Fanuc KAREL source: kt00743.KL

PROGRAM KT00743
%STACKSIZE=65535
%PRIORITY=65535
%NOLOCKGROUP
VAR
ARG : ARRAY[4] OF VECTOR
OUT : INTEGER
BEGIN
-- UNSAFE_SOURCE_IR line 7: OUT = native_s16_value(ARG)
END KT00743
